(* Schneider Machine Expert - Basic project Counter, file version 2.9.0.0 *)
(* ProjectInformations: Name=New project *)

HARDWARE
  Cpu 0: TM221M16R/G
  EthernetConfiguration: NetworkName=M221, IpAllocationMode=FixedAddress, IpAddress=0.0.0.0, SubnetMask=0.0.0.0
  SerialLineConfiguration: Baud=Baud19200, Parity=ParityEven, DataBits=DataBits8, StopBits=StopBits1, PhysicalMedium=PhysicalMediumRs485, TransmissionMode=TransmissionModeModbusRtu, SlaveId=1, Addressing=SlaveAddressing
  MastTask: UsePeriodScanMode=false, PeriodScan=100
  FastTask: Period=255
  CpuBehavior: StartingMode=StartAsPreviousState, AutoSaveRamOnEeprom=true, WatchdogPeriod=250

SYMBOLS  (address, symbol, comment, settings)
  %M0       A
  %M1       B
  %M3       C

POU New POU
  (* SectionNumber=1 *)

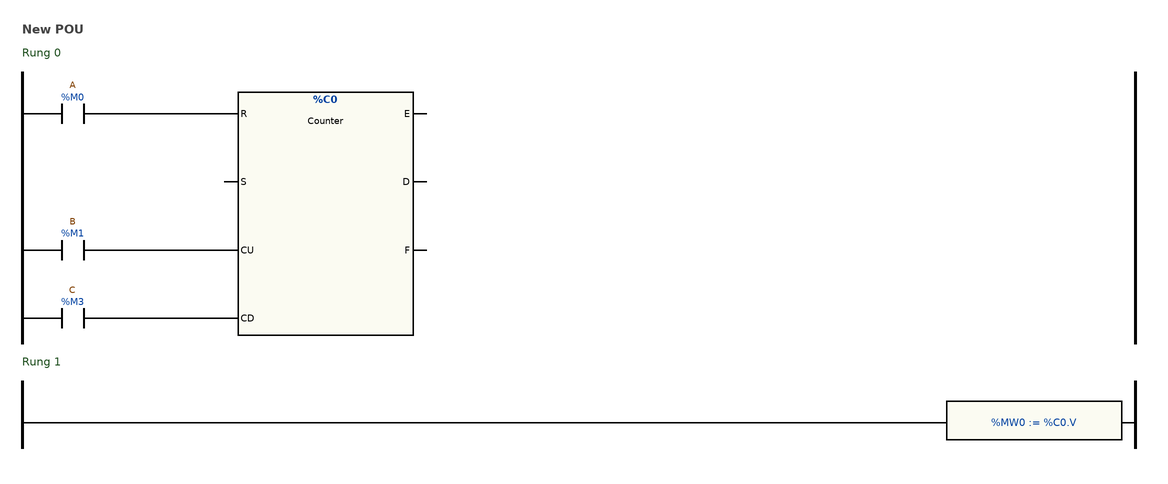

// Rung 0
  BLK %C0
  LD %M0                  (* A *)
  R
  LD %M1                  (* B *)
  CU
  LD %M3                  (* C *)
  CD
  END_BLK
  // as ST:
  //   %C0(R := A, CU := B, CD := C);

// Rung 1
  LD 1
  [ %MW0 := %C0.V ]
  // as ST:
  //   %MW0 := %C0.V;
